(* IEC 61131-3 sources: 2026_Projet_YGO_ExcavatriceDragage/CODE/J_SUPERVISION/_TYPES/8_BANDEAU_ET_IHM, 3 files *)

(* ---- ST_AlarmBanner.st ---- *)
(* ═══════════════════════════════════════════════════════════════
   🚨 ST_AlarmBanner — Bandeau d'alarme defilant (carrousel n/N)
   ───────────────────────────────────────────────────────────────
   🎯 Role : liste les defauts/warnings actifs de toute la machine,
      affiches un a la fois en rotation (FB_Hmi_BannerFormatter S5)
   📄 Doc : DOC/AF/AF_Partie-07_Interface_IHM_v2.3.md S6
   ═══════════════════════════════════════════════════════════════ *)
TYPE ST_AlarmBanner :
STRUCT
    HasAlarm    : BOOL;                        (* TRUE = au moins un defaut/warning actif *)
    Text        : STRING(120);                 (* Texte du message courant : [ORGANE] raison breve *)
    Index       : INT;                         (* Position courante (1-based, 0 si aucun defaut) *)
    Count       : INT;                         (* Nombre total de messages actifs *)
    AlarmArray  : ARRAY[0..49] OF STRING(120); (* 📋 Liste complete instantanee de tous les defauts actifs *)
END_STRUCT
END_TYPE

(* ---- ST_PermitVisibilityHMI.st ---- *)
(* Tableau public, lecture seule, des permis canoniques. Producteur : PRG_07. *)
TYPE ST_PermitVisibilityHMI :
STRUCT
    ArmingPermit : BOOL;
    M1SafetyAscentPermit : BOOL;
    M1SafetyDescendPermit : BOOL;
    M1ProcessAscentPermit : BOOL;
    M1ProcessDescendPermit : BOOL;
    EffectivePermitM1_Ascent : BOOL;
    EffectivePermitM1_Descend : BOOL;
    AppliedPermitM1_Ascent : BOOL;
    AppliedPermitM1_Descend : BOOL;
    M1FinalPermitBlocked : BOOL;
    M2SafetyAscentPermit : BOOL;
    M2SafetyDescendPermit : BOOL;
    M2ProcessAscentPermit : BOOL;
    M2ProcessDescendPermit : BOOL;
    EffectivePermitM2_Ascent : BOOL;
    EffectivePermitM2_Descend : BOOL;
    AppliedPermitM2_Ascent : BOOL;
    AppliedPermitM2_Descend : BOOL;
    M2FinalPermitBlocked : BOOL;
    BothActive : BOOL;
    BothBlocked : BOOL;
    BothBlockReason : E_WinchTraceBlockReason;
    EffectivePermitM3_Tremie : BOOL;
    EffectivePermitM3_Maintenance : BOOL; // Droit directionnel zone Maintenance, distinct de l'acces P1
    M3MotionPermitEffective : BOOL;
    DiveDescendPermit : BOOL;
    ExtractionAscentPermit : BOOL;
    ExtractionAssistActive : BOOL;
    EffectivePermitBucket_Open : BOOL;
    EffectivePermitBucket_Close : BOOL;
    // Benne : demandes et diagnostic d'execution, distincts des permis canoniques.
    BucketOpenRequestActive : BOOL;
    BucketCloseRequestActive : BOOL;
    BucketMotionBlocked : BOOL;
END_STRUCT
END_TYPE

(* ---- ST_PreflightHMI.st ---- *)
TYPE ST_PreflightHMI :
STRUCT
    BtnRun : BOOL;
    PreflightOk : BOOL;
    PreflightDone : BOOL;
    PreflightBusy : BOOL;
    PreflightErrorId : WORD;
END_STRUCT
END_TYPE
